FUNCTION_BLOCK Gerador_Generico (* Grupo gerador com DEIF AGC 150 - HidrycoLib *)
  (* Standard: 61499-2 *)
  (* Version 1.1, 15/10/2026, Hidryco, Hidryco, 1.1: comandos basicos da IHM (automatico, semiautomatico, partir e parar so em semiautomatico, reconhecer alarmes do AGC) nas palavras de comando 5 e 6 do AGC, publicadas em ${PATH}agcCmd5 e ${PATH}agcCmd6 (INT) para um MODBUSWREG2 no endereco 5; pulso de cfgTempoComando s, depois as palavras voltam a 0. 1.0: grupo gerador com controlador DEIF AGC 150 (aplicacao GEN, QTA com GB e MB). Leitura Modbus TCP FC04 pela configuracao de hardware (MODBUSGENTCPS + 9 MODBUSRREG8: 501, 513, 521, 536, 554, 567, 593, 1005, 1013); os registradores sao publicados nos symlinks ${PATH}rVAB ... ${PATH}rW1020 (INT) e o connStatusInt em ${PATH}comInt. Enderecos e escalas da tabela DEIF rev. S (software 1.19). *)
  PACKAGE Hidryco.HidrycoLib;
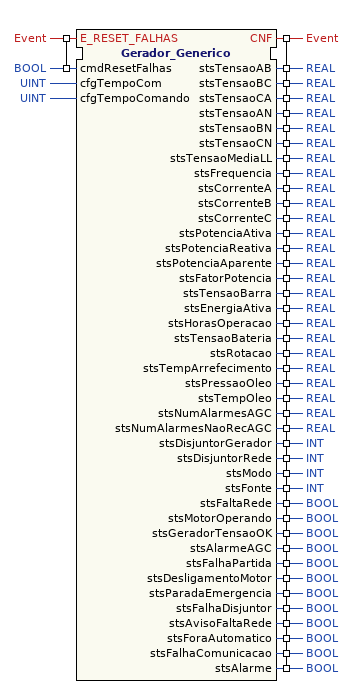
  EVENT_INPUT
    E_RESET_FALHAS WITH cmdResetFalhas; (* Reconhecimento pelo processo com cmdResetFalhas = TRUE *)
  END_EVENT
  EVENT_OUTPUT
    CNF WITH stsTensaoAB, stsTensaoBC, stsTensaoCA, stsTensaoAN, stsTensaoBN, stsTensaoCN, stsTensaoMediaLL, stsFrequencia, stsCorrenteA, stsCorrenteB, stsCorrenteC, stsPotenciaAtiva, stsPotenciaReativa, stsPotenciaAparente, stsFatorPotencia, stsTensaoBarra, stsEnergiaAtiva, stsHorasOperacao, stsTensaoBateria, stsRotacao, stsTempArrefecimento, stsPressaoOleo, stsTempOleo, stsNumAlarmesAGC, stsNumAlarmesNaoRecAGC, stsDisjuntorGerador, stsDisjuntorRede, stsModo, stsFonte, stsFaltaRede, stsMotorOperando, stsGeradorTensaoOK, stsAlarmeAGC, stsFalhaPartida, stsDesligamentoMotor, stsParadaEmergencia, stsFalhaDisjuntor, stsAvisoFaltaRede, stsForaAutomatico, stsFalhaComunicacao, stsAlarme; (* Valores e estados (so na mudanca) *)
  END_EVENT
  VAR_INPUT
    cmdResetFalhas : BOOL; (* TRUE = reconhecimento (com o evento E_RESET_FALHAS) *)
    cfgTempoCom : UINT := 10; (* Tempo (s) sem comunicacao com o AGC 150 para confirmar a falha *)
    cfgTempoComando : UINT := 2; (* Tempo (s) que a palavra de comando fica escrita no AGC *)
  END_VAR
  VAR_OUTPUT
    stsTensaoAB : REAL; (* Tensao A-B (V) *)
    stsTensaoBC : REAL; (* Tensao B-C (V) *)
    stsTensaoCA : REAL; (* Tensao C-A (V) *)
    stsTensaoAN : REAL; (* Tensao A-N (V) *)
    stsTensaoBN : REAL; (* Tensao B-N (V) *)
    stsTensaoCN : REAL; (* Tensao C-N (V) *)
    stsTensaoMediaLL : REAL; (* Tensao media fase-fase (V) *)
    stsFrequencia : REAL; (* Frequencia (Hz) *)
    stsCorrenteA : REAL; (* Corrente fase A (A) *)
    stsCorrenteB : REAL; (* Corrente fase B (A) *)
    stsCorrenteC : REAL; (* Corrente fase C (A) *)
    stsPotenciaAtiva : REAL; (* Potencia ativa (kW) *)
    stsPotenciaReativa : REAL; (* Potencia reativa (kVAr) *)
    stsPotenciaAparente : REAL; (* Potencia aparente (kVA) *)
    stsFatorPotencia : REAL; (* Fator de potencia *)
    stsTensaoBarra : REAL; (* Tensao do lado B (barramento/rede) L1-L2 (V) *)
    stsEnergiaAtiva : REAL; (* Energia ativa exportada (kWh) *)
    stsHorasOperacao : REAL; (* Horas de funcionamento (h) *)
    stsTensaoBateria : REAL; (* Tensao da bateria (V) *)
    stsRotacao : REAL; (* Rotacao do motor (rpm) *)
    stsTempArrefecimento : REAL; (* Temperatura do liquido de arrefecimento (°C) *)
    stsPressaoOleo : REAL; (* Pressao do oleo (bar) *)
    stsTempOleo : REAL; (* Temperatura do oleo (°C) *)
    stsNumAlarmesAGC : REAL; (* Alarmes ativos no AGC *)
    stsNumAlarmesNaoRecAGC : REAL; (* Alarmes nao reconhecidos no AGC *)
    stsDisjuntorGerador : INT; (* Disjuntor do gerador (GB): 0 indefinido/sem comunicacao, 1 aberto, 2 fechado *)
    stsDisjuntorRede : INT; (* Disjuntor de rede (MB): 0 indefinido/sem comunicacao, 1 aberto, 2 fechado *)
    stsModo : INT; (* Modo do AGC: 0 indefinido, 1 automatico, 2 semi-automatico, 3 manual, 4 bloqueio, 5 teste *)
    stsFonte : INT; (* Fonte da saida do QTA: 0 sem fonte, 1 rede, 2 gerador, 3 indefinida (sem comunicacao) *)
    stsFaltaRede : BOOL; (* Falta de rede (AMF) *)
    stsMotorOperando : BOOL; (* Motor em operacao *)
    stsGeradorTensaoOK : BOOL; (* Tensao e frequencia do gerador OK *)
    stsAlarmeAGC : BOOL; (* Alarme ativo no controlador do gerador (AGC 150) *)
    stsFalhaPartida : BOOL; (* Falha na partida do gerador *)
    stsDesligamentoMotor : BOOL; (* Desligamento do motor (ECU ou sobrevelocidade) *)
    stsParadaEmergencia : BOOL; (* Parada de emergência do gerador acionada *)
    stsFalhaDisjuntor : BOOL; (* Falha de disjuntor no QTA (gerador ou rede) *)
    stsAvisoFaltaRede : BOOL; (* Falta de rede no QTA *)
    stsForaAutomatico : BOOL; (* Gerador fora do modo automático *)
    stsFalhaComunicacao : BOOL; (* Falha de comunicacao com o AGC 150 *)
    stsAlarme : BOOL; (* Algum alarme do gerador *)
  END_VAR
  FBS
    IThis : Gerador_Generico_HMI(QI := TRUE);
    plcStart1 : plcStart(Prio := 10);
    Logica : basicGeradorGenerico;
    Tick : E_CYCLE(DT := T#1s);
    Leitura1 : SYMLINKMULTIVARDST_115C998103CD7017B(NAME1 := '$${PATH}rVAB', NAME2 := '$${PATH}rVBC', NAME3 := '$${PATH}rVCA', NAME4 := '$${PATH}rVAN', NAME5 := '$${PATH}rVBN', NAME6 := '$${PATH}rVCN', NAME7 := '$${PATH}rFreq', NAME8 := '$${PATH}rIA', NAME9 := '$${PATH}rIB', NAME10 := '$${PATH}rIC', NAME11 := '$${PATH}rPAtiva', NAME12 := '$${PATH}rQReativa', NAME13 := '$${PATH}rSAparente', NAME14 := '$${PATH}rFP', NAME15 := '$${PATH}rVBarra', QI := TRUE); {SET_ATTRIBUTE(Configuration.GenericFBType.InterfaceParams, Runtime.System#I:=15;VALUE${I$}:INT,INT,INT,INT,INT,INT,INT,INT,INT,INT,INT,INT,INT,INT,INT)}
    Leitura2 : SYMLINKMULTIVARDST_115C998103CD7017B(NAME1 := '$${PATH}rEnergiaH', NAME2 := '$${PATH}rEnergiaL', NAME3 := '$${PATH}rHorasH', NAME4 := '$${PATH}rHorasL', NAME5 := '$${PATH}rNumAlm', NAME6 := '$${PATH}rNumAlmNR', NAME7 := '$${PATH}rBateria', NAME8 := '$${PATH}rRPM', NAME9 := '$${PATH}rTempAgua', NAME10 := '$${PATH}rPressOleo', NAME11 := '$${PATH}rTempOleo', NAME12 := '$${PATH}rW1005', NAME13 := '$${PATH}rW1010', NAME14 := '$${PATH}rW1013', NAME15 := '$${PATH}rW1014', QI := TRUE); {SET_ATTRIBUTE(Configuration.GenericFBType.InterfaceParams, Runtime.System#I:=15;VALUE${I$}:INT,INT,INT,INT,INT,INT,INT,INT,INT,INT,INT,INT,INT,INT,INT)}
    Leitura3 : SYMLINKMULTIVARDST_15292F208F22048C1(NAME1 := '$${PATH}rW1015', NAME2 := '$${PATH}rW1018', NAME3 := '$${PATH}rW1019', NAME4 := '$${PATH}rW1020', QI := TRUE); {SET_ATTRIBUTE(Configuration.GenericFBType.InterfaceParams, Runtime.System#I:=4;VALUE${I$}:INT,INT,INT,INT)}
    Comunicacao : SYMLINKMULTIVARDST_5A03F112CD5D470(NAME1 := '$${PATH}comInt', QI := TRUE); {SET_ATTRIBUTE(Configuration.GenericFBType.InterfaceParams, Runtime.System#I:=1;VALUE${I$}:INT)}
    AlarmeAGC : ALARM_BIT(TYPE := 1, ACKTYPE_1 := 2, ACTIVE := TRUE); {SET_ATTRIBUTE(HMI.AlarmText, Alarme ativo no controlador do gerador (AGC 150))}
    AlarmePartida : ALARM_BIT(TYPE := 1, ACKTYPE_1 := 2, ACTIVE := TRUE); {SET_ATTRIBUTE(HMI.AlarmText, Falha na partida do gerador)}
    AlarmeMotor : ALARM_BIT(TYPE := 1, ACKTYPE_1 := 2, ACTIVE := TRUE); {SET_ATTRIBUTE(HMI.AlarmText, Motor do gerador desligado por proteção (ECU ou sobrevelocidade))}
    AlarmeEmergencia : ALARM_BIT(TYPE := 1, ACKTYPE_1 := 2, ACTIVE := TRUE); {SET_ATTRIBUTE(HMI.AlarmText, Parada de emergência do gerador acionada)}
    AlarmeDisjuntor : ALARM_BIT(TYPE := 1, ACKTYPE_1 := 2, ACTIVE := TRUE); {SET_ATTRIBUTE(HMI.AlarmText, Falha de disjuntor no QTA (gerador ou rede))}
    AlarmeFaltaRede : ALARM_BIT(TYPE := 1, ACKTYPE_1 := 2, ACTIVE := TRUE); {SET_ATTRIBUTE(HMI.AlarmText, Falta de energia da rede no QTA)} {SET_ATTRIBUTE(HMI.AlarmClass, Warning)}
    AlarmeForaAuto : ALARM_BIT(TYPE := 1, ACKTYPE_1 := 2, ACTIVE := TRUE); {SET_ATTRIBUTE(HMI.AlarmText, Gerador fora do modo automático)} {SET_ATTRIBUTE(HMI.AlarmClass, Warning)}
    AlarmeComunicacao : ALARM_BIT(TYPE := 1, ACKTYPE_1 := 2, ACTIVE := TRUE); {SET_ATTRIBUTE(HMI.AlarmText, Controlador do gerador (AGC 150) sem comunicação)}
    ComandoAGC5 : SYMLINKMULTIVARSRC_5A03F112CD5D470(NAME1 := '$${PATH}agcCmd5', QI := TRUE); {SET_ATTRIBUTE(Configuration.GenericFBType.InterfaceParams, Runtime.System#I:=1;VALUE${I$}:INT)}
    ComandoAGC6 : SYMLINKMULTIVARSRC_5A03F112CD5D470(NAME1 := '$${PATH}agcCmd6', QI := TRUE); {SET_ATTRIBUTE(Configuration.GenericFBType.InterfaceParams, Runtime.System#I:=1;VALUE${I$}:INT)}
  END_FBS
  EVENT_CONNECTIONS
    plcStart1.FIRST_INIT TO IThis.E97FC986B98F8068;
    plcStart1.REDO_INIT TO IThis.E97FC986B98F8068;
    IThis.E947B6720B0429AC TO Logica.2BF6A84D5AF65FB4;
    Logica.DC12539614B57B73 TO Tick.START;
    Logica.DC12539614B57B73 TO Leitura1.INIT;
    Logica.DC12539614B57B73 TO Leitura2.INIT;
    Logica.DC12539614B57B73 TO Leitura3.INIT;
    Logica.DC12539614B57B73 TO Comunicacao.INIT;
    Logica.DC12539614B57B73 TO AlarmeAGC.INIT;
    AlarmeAGC.INITO TO AlarmeAGC.REQ_INITDATA;
    AlarmeAGC.CNF_INITDATA TO AlarmeAGC.ACTIVATE;
    AlarmeAGC.INITO TO AlarmePartida.INIT;
    AlarmePartida.INITO TO AlarmePartida.REQ_INITDATA;
    AlarmePartida.CNF_INITDATA TO AlarmePartida.ACTIVATE;
    AlarmePartida.INITO TO AlarmeMotor.INIT;
    AlarmeMotor.INITO TO AlarmeMotor.REQ_INITDATA;
    AlarmeMotor.CNF_INITDATA TO AlarmeMotor.ACTIVATE;
    AlarmeMotor.INITO TO AlarmeEmergencia.INIT;
    AlarmeEmergencia.INITO TO AlarmeEmergencia.REQ_INITDATA;
    AlarmeEmergencia.CNF_INITDATA TO AlarmeEmergencia.ACTIVATE;
    AlarmeEmergencia.INITO TO AlarmeDisjuntor.INIT;
    AlarmeDisjuntor.INITO TO AlarmeDisjuntor.REQ_INITDATA;
    AlarmeDisjuntor.CNF_INITDATA TO AlarmeDisjuntor.ACTIVATE;
    AlarmeDisjuntor.INITO TO AlarmeFaltaRede.INIT;
    AlarmeFaltaRede.INITO TO AlarmeFaltaRede.REQ_INITDATA;
    AlarmeFaltaRede.CNF_INITDATA TO AlarmeFaltaRede.ACTIVATE;
    AlarmeFaltaRede.INITO TO AlarmeForaAuto.INIT;
    AlarmeForaAuto.INITO TO AlarmeForaAuto.REQ_INITDATA;
    AlarmeForaAuto.CNF_INITDATA TO AlarmeForaAuto.ACTIVATE;
    AlarmeForaAuto.INITO TO AlarmeComunicacao.INIT;
    AlarmeComunicacao.INITO TO AlarmeComunicacao.REQ_INITDATA;
    AlarmeComunicacao.CNF_INITDATA TO AlarmeComunicacao.ACTIVATE;
    AlarmeComunicacao.INITO TO plcStart1.ACK_FIRST;
    Logica.DC12539614B57B73 TO ComandoAGC5.INIT;
    Logica.DC12539614B57B73 TO ComandoAGC6.INIT;
    Logica.C9337F6B69351BCF TO ComandoAGC5.REQ;
    Logica.C9337F6B69351BCF TO ComandoAGC6.REQ;
    IThis.6D578F9B82E559A7 TO Logica.15D59D6E025E0AEC;
    IThis.E92041950CEDCF19 TO Logica.D7C528B832D24695;
    E_RESET_FALHAS TO Logica.58BFBDBCB72060FA;
    Tick.EO TO Logica.1DB3A43D9CFE56D9;
    Logica.A44CBE1A3706F856 TO CNF;
    Logica.E2CCA36837A78D9A TO IThis.26D8CC00FA2A4527;
    Leitura1.CNF TO Logica.BDA6F58D663AD593;
    Leitura2.CNF TO Logica.11A3A648381739C8;
    Leitura3.CNF TO Logica.748B4B0803385F35;
    Comunicacao.CNF TO Logica.A19EF8FB897BEE21;
    Logica.0972B515C8BC4FF5 TO AlarmeAGC.REQ;
    Logica.0972B515C8BC4FF5 TO AlarmePartida.REQ;
    Logica.0972B515C8BC4FF5 TO AlarmeMotor.REQ;
    Logica.0972B515C8BC4FF5 TO AlarmeEmergencia.REQ;
    Logica.0972B515C8BC4FF5 TO AlarmeDisjuntor.REQ;
    Logica.0972B515C8BC4FF5 TO AlarmeFaltaRede.REQ;
    Logica.0972B515C8BC4FF5 TO AlarmeForaAuto.REQ;
    Logica.0972B515C8BC4FF5 TO AlarmeComunicacao.REQ;
    AlarmeAGC.IND_1 TO IThis.26D8CC00FA2A4527;
    AlarmePartida.IND_1 TO IThis.26D8CC00FA2A4527;
    AlarmeMotor.IND_1 TO IThis.26D8CC00FA2A4527;
    AlarmeEmergencia.IND_1 TO IThis.26D8CC00FA2A4527;
    AlarmeDisjuntor.IND_1 TO IThis.26D8CC00FA2A4527;
    AlarmeFaltaRede.IND_1 TO IThis.26D8CC00FA2A4527;
    AlarmeForaAuto.IND_1 TO IThis.26D8CC00FA2A4527;
    AlarmeComunicacao.IND_1 TO IThis.26D8CC00FA2A4527;
    IThis.E92041950CEDCF19 TO AlarmeAGC.ACK_C1;
    IThis.E92041950CEDCF19 TO AlarmePartida.ACK_C1;
    IThis.E92041950CEDCF19 TO AlarmeMotor.ACK_C1;
    IThis.E92041950CEDCF19 TO AlarmeEmergencia.ACK_C1;
    IThis.E92041950CEDCF19 TO AlarmeDisjuntor.ACK_C1;
    IThis.E92041950CEDCF19 TO AlarmeFaltaRede.ACK_C1;
    IThis.E92041950CEDCF19 TO AlarmeForaAuto.ACK_C1;
    IThis.E92041950CEDCF19 TO AlarmeComunicacao.ACK_C1;
    E_RESET_FALHAS TO AlarmeAGC.ACK_C1;
    E_RESET_FALHAS TO AlarmePartida.ACK_C1;
    E_RESET_FALHAS TO AlarmeMotor.ACK_C1;
    E_RESET_FALHAS TO AlarmeEmergencia.ACK_C1;
    E_RESET_FALHAS TO AlarmeDisjuntor.ACK_C1;
    E_RESET_FALHAS TO AlarmeFaltaRede.ACK_C1;
    E_RESET_FALHAS TO AlarmeForaAuto.ACK_C1;
    E_RESET_FALHAS TO AlarmeComunicacao.ACK_C1;
  END_CONNECTIONS
  DATA_CONNECTIONS
    cfgTempoCom TO Logica.5D2B8D5EEA8CA438;
    cfgTempoComando TO Logica.CBB484B85F481F97;
    cmdResetFalhas TO Logica.0D423F13A9758F5D;
    Leitura1.VALUE1 TO Logica.A7330B3B6EB1E31F;
    Leitura1.VALUE2 TO Logica.75CBA331281D5001;
    Leitura1.VALUE3 TO Logica.66EF7D2E67C68200;
    Leitura1.VALUE4 TO Logica.9C5E7398418C1F4F;
    Leitura1.VALUE5 TO Logica.EF4B3D706C982888;
    Leitura1.VALUE6 TO Logica.31E01BD221C0A7DE;
    Leitura1.VALUE7 TO Logica.245118D9851C76BB;
    Leitura1.VALUE8 TO Logica.FC48B87CE94C8360;
    Leitura1.VALUE9 TO Logica.13929E799CB18846;
    Leitura1.VALUE10 TO Logica.AAC42DE962D3B797;
    Leitura1.VALUE11 TO Logica.2B4EE563F848EAD2;
    Leitura1.VALUE12 TO Logica.D9530A834C71219B;
    Leitura1.VALUE13 TO Logica.61A9D188A9F5851B;
    Leitura1.VALUE14 TO Logica.5C1EE40821C23758;
    Leitura1.VALUE15 TO Logica.982869116272FA7B;
    Leitura2.VALUE1 TO Logica.D7521402DC916D5E;
    Leitura2.VALUE2 TO Logica.F9EA42AE519A3D2E;
    Leitura2.VALUE3 TO Logica.63486372C36DDBF8;
    Leitura2.VALUE4 TO Logica.F4ABDF0B282740AC;
    Leitura2.VALUE5 TO Logica.EBAD8D198B0E57E2;
    Leitura2.VALUE6 TO Logica.0BADCB814AA024F4;
    Leitura2.VALUE7 TO Logica.DC4211A23853BF02;
    Leitura2.VALUE8 TO Logica.021B316D2E9FC503;
    Leitura2.VALUE9 TO Logica.D0280F27AA894985;
    Leitura2.VALUE10 TO Logica.022589950134A15C;
    Leitura2.VALUE11 TO Logica.1D7067E42F7F920B;
    Leitura2.VALUE12 TO Logica.28086F9A13C4AEC8;
    Leitura2.VALUE13 TO Logica.B744057DFF29435F;
    Leitura2.VALUE14 TO Logica.E7BDF46B90F2ABE7;
    Leitura2.VALUE15 TO Logica.85B76D64ED703E5C;
    Leitura3.VALUE1 TO Logica.0B6F0F6CAFB73D0B;
    Leitura3.VALUE2 TO Logica.C0ECE3FD244E9D27;
    Leitura3.VALUE3 TO Logica.485CC684071F672F;
    Leitura3.VALUE4 TO Logica.49ACB6AFF371591F;
    Comunicacao.VALUE1 TO Logica.31128805057AE6DF;
    IThis.853136B9D18CF5B5 TO Logica.C2183108F3905F97;
    IThis.B1D3FD444B829FE6 TO Logica.7160EE4A63D00A51;
    Logica.2ACC4459D225B2A5 TO ComandoAGC5.VALUE1;
    Logica.600857C82B1F69BA TO ComandoAGC6.VALUE1;
    Logica.7282D542BDBB3FFB TO AlarmeAGC.INP;
    Logica.613FBFDAE9BD92D2 TO AlarmePartida.INP;
    Logica.F735731CEC5837CB TO AlarmeMotor.INP;
    Logica.3E0F2ACB4615C726 TO AlarmeEmergencia.INP;
    Logica.CE665728889A4341 TO AlarmeDisjuntor.INP;
    Logica.422AAB54CD83B326 TO AlarmeFaltaRede.INP;
    Logica.39057C2ACBA9565F TO AlarmeForaAuto.INP;
    Logica.91DD86BE95DDFBA8 TO AlarmeComunicacao.INP;
    Logica.1E40D0D699DD144E TO stsTensaoAB;
    Logica.C19F83948281B0E2 TO stsTensaoBC;
    Logica.3C88756B36A52512 TO stsTensaoCA;
    Logica.4BA5F5355FF4CEA7 TO stsTensaoAN;
    Logica.E36E8F1BEC8ADC88 TO stsTensaoBN;
    Logica.CA33BD0236498767 TO stsTensaoCN;
    Logica.F19F5E032DA269A0 TO stsTensaoMediaLL;
    Logica.B4ED2B665DF935CA TO stsFrequencia;
    Logica.224868A578BADC0A TO stsCorrenteA;
    Logica.C1F286943C35525A TO stsCorrenteB;
    Logica.3A87AFDA0837A305 TO stsCorrenteC;
    Logica.953A300991140BB0 TO stsPotenciaAtiva;
    Logica.7395FF5E7D3E1486 TO stsPotenciaReativa;
    Logica.CA2CF5BB08A1B5AC TO stsPotenciaAparente;
    Logica.95830401F9DB0E6C TO stsFatorPotencia;
    Logica.D05459853BFE584C TO stsTensaoBarra;
    Logica.80875DDED85C9768 TO stsEnergiaAtiva;
    Logica.42A342504DB52425 TO stsHorasOperacao;
    Logica.DD82132D7F9E0054 TO stsTensaoBateria;
    Logica.F2420F8AB10CFA35 TO stsRotacao;
    Logica.D14EBEC5B3C194C5 TO stsTempArrefecimento;
    Logica.0E8548B50BBA41D7 TO stsPressaoOleo;
    Logica.2053820AB993FCDC TO stsTempOleo;
    Logica.C733850F46B2B7C0 TO stsNumAlarmesAGC;
    Logica.51695C60F1D860CF TO stsNumAlarmesNaoRecAGC;
    Logica.39EB84F933B4E6D9 TO stsDisjuntorGerador;
    Logica.692FFC497509E0A1 TO stsDisjuntorRede;
    Logica.C084ABF0328A5376 TO stsModo;
    Logica.9172A58AE36C8C37 TO stsFonte;
    Logica.7F54324733CC63A1 TO stsFaltaRede;
    Logica.29A1CBB8F7435B76 TO stsMotorOperando;
    Logica.36CCB0EB6EDA1E16 TO stsGeradorTensaoOK;
    Logica.3FBFE0CD60124175 TO stsAlarmeAGC;
    Logica.60591644B144BF74 TO stsFalhaPartida;
    Logica.D0B870E4138B8E9A TO stsDesligamentoMotor;
    Logica.996A96555603652B TO stsParadaEmergencia;
    Logica.D6D6D24B3FBF0ADC TO stsFalhaDisjuntor;
    Logica.A7E5F1F016368C29 TO stsAvisoFaltaRede;
    Logica.F41F41A2F194D1F0 TO stsForaAutomatico;
    Logica.A4FF00541968E223 TO stsFalhaComunicacao;
    Logica.69B14C75210049E3 TO stsAlarme;
    Logica.1E40D0D699DD144E TO IThis.00413B77FB3FD391;
    Logica.C19F83948281B0E2 TO IThis.6FB2F6B28DC276BC;
    Logica.3C88756B36A52512 TO IThis.61ECA2065F4A1220;
    Logica.4BA5F5355FF4CEA7 TO IThis.C55D1A7D24318BE9;
    Logica.E36E8F1BEC8ADC88 TO IThis.B3C1C2B1D84A8BEF;
    Logica.CA33BD0236498767 TO IThis.A9BCCDA5C9491BC5;
    Logica.F19F5E032DA269A0 TO IThis.6D6FCE7EEF5A092F;
    Logica.B4ED2B665DF935CA TO IThis.A6B15948115E4622;
    Logica.224868A578BADC0A TO IThis.06755BC431017794;
    Logica.C1F286943C35525A TO IThis.48E59B4224572852;
    Logica.3A87AFDA0837A305 TO IThis.546F39FA179BDCFE;
    Logica.953A300991140BB0 TO IThis.D45ADC0A6454CCC7;
    Logica.7395FF5E7D3E1486 TO IThis.C25D419DB7DBCFF4;
    Logica.CA2CF5BB08A1B5AC TO IThis.5DD3E088782C8D1B;
    Logica.95830401F9DB0E6C TO IThis.DC02F918C07495F6;
    Logica.D05459853BFE584C TO IThis.B15E2E9E8D19A37F;
    Logica.80875DDED85C9768 TO IThis.843AFFBDAD6A0A35;
    Logica.42A342504DB52425 TO IThis.D96330EF0A6E3612;
    Logica.DD82132D7F9E0054 TO IThis.4C9948807F71F264;
    Logica.F2420F8AB10CFA35 TO IThis.226B306D451A97EB;
    Logica.D14EBEC5B3C194C5 TO IThis.21DCDE8193E3FBEF;
    Logica.0E8548B50BBA41D7 TO IThis.B9558F209B183E4E;
    Logica.2053820AB993FCDC TO IThis.7E4E6F21D9F3B7B2;
    Logica.C733850F46B2B7C0 TO IThis.544D9AC77812BDA1;
    Logica.51695C60F1D860CF TO IThis.646698EA651C1295;
    Logica.39EB84F933B4E6D9 TO IThis.0C2444BAA28C89B4;
    Logica.692FFC497509E0A1 TO IThis.3FCEB32B27865B69;
    Logica.C084ABF0328A5376 TO IThis.7138AB6343D50B72;
    Logica.9172A58AE36C8C37 TO IThis.5B3A9F4868BF85D1;
    Logica.7F54324733CC63A1 TO IThis.9ADF793C78EB9815;
    Logica.29A1CBB8F7435B76 TO IThis.040C3BE2C9BFF722;
    Logica.36CCB0EB6EDA1E16 TO IThis.E94B12BF1E46D1DE;
    Logica.3FBFE0CD60124175 TO IThis.8DFB812BDDFA5844;
    Logica.60591644B144BF74 TO IThis.3C3153BF8E08E275;
    Logica.D0B870E4138B8E9A TO IThis.D0DBD7A32CDF5CF0;
    Logica.996A96555603652B TO IThis.AC299F89EBF46FB1;
    Logica.D6D6D24B3FBF0ADC TO IThis.7509DCD3B4E54882;
    Logica.A7E5F1F016368C29 TO IThis.B935E662D3F620E5;
    Logica.F41F41A2F194D1F0 TO IThis.E9CE0A38EB06D84D;
    Logica.A4FF00541968E223 TO IThis.F9C5A53F446008C4;
    Logica.69B14C75210049E3 TO IThis.BDC6AA03EB5CCBEC;
    AlarmeAGC.STATE_1 TO IThis.A40DB40432E241B0;
    AlarmePartida.STATE_1 TO IThis.4D16197CC8A6FA3A;
    AlarmeMotor.STATE_1 TO IThis.B623E8D435377242;
    AlarmeEmergencia.STATE_1 TO IThis.AF8683B23D9C1DA8;
    AlarmeDisjuntor.STATE_1 TO IThis.34A389507308939C;
    AlarmeFaltaRede.STATE_1 TO IThis.D79A25D4A4B48D7C;
    AlarmeForaAuto.STATE_1 TO IThis.E9D8329650B83C14;
    AlarmeComunicacao.STATE_1 TO IThis.00731EA1F129697D;
    Logica.C2B751B97236C67C TO IThis.D970C941743E38D2;
    Logica.3A929C8EED3B371D TO IThis.0B3DF6FBECF5CB74;
    Logica.840FF50E52A3339F TO IThis.ED00303F35471587;
    Logica.0D4A3E26781F6D90 TO IThis.BB32D518A4DF7385;
    Logica.EFA6B10159DC226B TO IThis.E4D7528507F03FF0;
    Logica.3A1C7F4B518A0AFA TO IThis.3A49104F51FAE798;
  END_CONNECTIONS
END_FUNCTION_BLOCK
